RESOURCE RES0 : EMB_RES_ECO
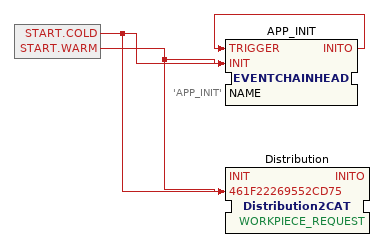
  FBS
    Distribution : Distribution2CAT;
    APP_INIT : EVENTCHAINHEAD(NAME := 'APP_INIT');
  END_FBS
  EVENT_CONNECTIONS
    APP_INIT.INITO TO APP_INIT.TRIGGER;
    START.COLD TO Distribution.461F22269552CD75;
    START.WARM TO Distribution.461F22269552CD75;
    START.COLD TO APP_INIT.INIT;
    START.WARM TO APP_INIT.INIT;
  END_CONNECTIONS
END_RESOURCE
